// TIA Portal V21 export
// export: Created 2026-08-21T20:18:56.5189349Z, ExportSetting None, DisplayName Totally Integrated Automation Portal, DisplayVersion V21, DisplayName STEP 7 Professional, DisplayVersion V21, DisplayName STEP 7 Safety, DisplayVersion V21, DisplayName Tech WebApplication, DisplayVersion V21, DisplayName WinCC Basic/Comfort/Advanced, DisplayVersion V21, DisplayName WinCC Professional, DisplayVersion V21, DisplayName WinCC Unified, DisplayVersion V21
TYPE "UDT_Service_StatusMedium"
   STRUCT
      parameterError { ExternalWritable := 'False'} : Bool := FALSE;   // ParameterStart & ParameterEnd area out of range
      parameterTypeError { ExternalWritable := 'False'} : Bool;   // Parametertype not defined; Number of Type out of range
      monitoringTimeExceeded { ExternalWritable := 'False'} : Bool := FALSE;   // Step monitoring time exceeded
      noSystemTime { ExternalWritable := 'False'} : Bool;   // FB cannot evaluate system / sample time
      SteporderStatus { ExternalWritable := 'False'} : Array[0..6] of DWord;   // Indication of steporder state
   END_STRUCT;
END_TYPE
